FUNCTION_BLOCK basicStatusRemota (* Estado da comunicacao de uma remota Modbus TCP *)
  (* Standard: 61499-2 *)
  (* Version 1.1, 06/11/2026, Hidryco, Hidryco, 1.1: aceita 'Online' (valor real do runtime; antes so 'online' e toda remota comunicando aparecia SEM COMUNICACAO); INIT tambem le o conn (antes o valor inicial era ignorado e a remota ficava AGUARDANDO); CNF_HMI a cada leitura com stsVivo (sinal de vida para a IHM). 1.0: connStatus (online/offline) do escravo MODBUSGENTCPS *)
  PACKAGE Hidryco.HidrycoLib;
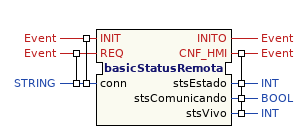
  EVENT_INPUT
    INIT WITH conn; (* Inicializacao (com o valor atual do connStatus) *)
    REQ WITH conn; (* Status da conexao recebido do hardware *)
  END_EVENT
  EVENT_OUTPUT
    INITO; (* Inicializacao concluida *)
    CNF_HMI WITH stsEstado, stsComunicando, stsVivo; (* Status para a IHM (a cada leitura) *)
  END_EVENT
  VAR_INPUT
    conn : STRING; (* connStatus do escravo Modbus TCP: online / offline *)
  END_VAR
  VAR_OUTPUT
    stsEstado : INT; (* 0 aguardando, 1 comunicando, 2 sem comunicacao *)
    stsComunicando : BOOL; (* Remota comunicando *)
    stsVivo : INT; (* Sinal de vida: contador 0..9999 a cada leitura *)
  END_VAR
  VAR
    initDone : BOOL;
    primeiro : BOOL := TRUE;
    est : INT;
    oldEst : INT := -1;
    vivo : INT;
  END_VAR
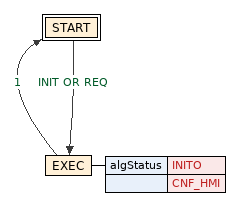
  EC_STATES
    START; (* Estado inicial *)
    EXEC : algStatus -> INITO, -> CNF_HMI; (* Executa a logica; o algoritmo decide quais eventos saem *)
  END_STATES
  EC_TRANSITIONS
    START TO EXEC := INIT OR REQ;
    EXEC TO START := 1;
  END_TRANSITIONS
  ALGORITHM algStatus IN ST: (* Logica completa *)
(* =====================================================================
   basicStatusRemota v1.1 - estado da comunicacao de uma remota
   connStatus do MODBUSGENTCPS: o runtime manda 'Online' / 'Offline' (conferido online no EAE 06/11/2026;
   a documentacao diz 'online'): aceita as tres grafias.
   INIT tambem le o conn (valor atual entregue no INITO do symlink).
   Cada INIT/REQ emite CNF_HMI com stsVivo (contador) para a IHM detectar CLP sem dados.
   ===================================================================== *)
INITO   := FALSE;
CNF_HMI := FALSE;
IF INIT THEN
    initDone := TRUE;
    INITO := TRUE;
END_IF;
IF NOT initDone THEN
    RETURN;
END_IF;
IF (conn = 'Online') OR (conn = 'online') OR (conn = 'ONLINE') THEN
    est := 1;
ELSIF conn = '' THEN
    est := 0;
ELSE
    est := 2;
END_IF;
stsEstado := est;
stsComunicando := est = 1;
vivo := vivo + 1;
IF vivo > 9999 THEN
    vivo := 0;
END_IF;
stsVivo := vivo;
CNF_HMI := TRUE;
  END_ALGORITHM
END_FUNCTION_BLOCK
